(* IEC 61131-3 sources: Elmo_Master/Lasal_PRG/Elmo_EtherCAT_Test_4Axis/Class/CP733_IOs, 1 file *)

(* ---- CP733_IOs.st ---- *)
//FPGA Components
#define CP733_IOS_DEVICE_ID_XADC           16#0A60
#define CP733_IOS_DEVICE_ID_CPU_REG        16#0F02

//XADC Register
#define CP733_IOS_OFFSET_TEMPERATURE       16#00
#define CP733_IOS_OFFSET_VOLTAGE_VP_VN     16#06
#define CP733_IOS_OFFSET_TEMPERATURE_MAX   16#40
#define CP733_IOS_OFFSET_TEMPERATURE_MIN   16#48

//CPU Register
#define CP733_IOS_OFFSET_DIGITAL_INPUT_REGISTER           16#00
#define CP733_IOS_OFFSET_DIGITAL_OUTPUT_CLEAR_REGISTER    16#01
#define CP733_IOS_OFFSET_DIGITAL_OUTPUT_READ_SET_REGISTER 16#02

#define CP733_IOS_REGISTER_NOT_FOUND       16#FFFF

#define CP733_IOS_OFFSET_TEMPSENSOR1       16#08
#define CP733_IOS_OFFSET_TEMPSENSOR2       16#0A

//Constants and calculation from xilinx datasheet
//https://www.xilinx.com/support/documentation/user_guides/ug480_7Series_XADC.pdf
//Equation 2-6 (Temperature) and Equation 2-7 (Voltage)
#define CP733_TEMP_MULTIPLIER    503.975
#define CP733_TEMP_DIVISIOR      4096
#define CP733_TEMP_OFFSET        273.15

#define CP733_IOS_TEMP_CONSTANT_KELVIN  273

#define CP733_VOLTAGE_MULTIPLIER 31

#define CP733_CONVERT_V_TO_MV    1000    //Convert V to mV
#define CP733_CONVERT_TO_1_10_C  10      //Convert °C to 1/10 °C

#define CP733_SUPPLY_VOLTAGE_OFFSET 430  //0,43 V offset (Info from CPU department)

#include "..\..\Source\interfaces\lsl_st_pci.h"
#include "..\..\Source\interfaces\lsl_st_xadc.h"
#include "..\..\Class\PLC_Info\XRegs.h"
#include "..\..\Source\interfaces\lsl_st_gpio.h"

(*!
<Class
	Name               = "CP733_IOs"
	Revision           = "1.0"
	RealtimeTask       = "false"
	CyclicTask         = "false"
	BackgroundTask     = "false"
	Sigmatek           = "true"
	OSInterface        = "false"
	HighPriority       = "false"
	Automatic          = "false"
	UpdateMode         = "Prescan"
	IconPath           = ".\Class\DigInOut.ICO"
	SharedCommandTable = "true"
	Objectsize         = "(688,120)"
	Comment            = "Hardwareclass to access the IOs on the CP733.">
	<Channels>
		<Server Name="BatteryOk" Visualized="true" Initialize="false" WriteProtected="true" Retentive="false" Comment="Shows the state of the battery.&#13;&#10;0 .. Not OK&#13;&#10;1 .. OK"/>
		<Server Name="Can1_Termination" Visualized="true" Initialize="true" WriteProtected="false" Retentive="false" Comment="Write to this server to set the CAN termination.&#13;&#10;0 ... CAN termination is off&#13;&#10;1 ... CAN termination is on&#13;&#10;-1 ... not available/failed to set register in FPGA"/>
		<Server Name="CAN_1_Connect" Class="_CanLib" Visualized="false" Initialize="false" WriteProtected="true" Retentive="false"/>
		<Server Name="ClassState" Visualized="true" Initialize="false" WriteProtected="true" Retentive="false" Comment="Shows the initialisation state of the class.&#13;&#10; 0 ... Initialisation ok&#13;&#10;-1 ... PCI Interface not found&#13;&#10;-2 ... &quot;XADC&quot; interface not found&#13;&#10;-3 ... &quot;IXREGS&quot; interface not found&#13;&#10;-4 ... GPIO Interface not found&#13;&#10;-5 ... CPU Register not found&#13;&#10;-6 ... Login to HwControl failed&#13;&#10;"/>
		<Server Name="ErrorLED" Visualized="true" Initialize="false" WriteProtected="false" Retentive="false" Comment="The &quot;Error&quot;-LED of the CPU can be controlled with this server.&#13;&#10;&#13;&#10;0 ... HW - Status of LED is active&#13;&#10;1 ... LED is off&#13;&#10;2 ... LED is flashes&#13;&#10;3 ... LED is on&#13;&#10;&#13;&#10;-1 ... Class not ok"/>
		<Server Name="Ethernet_1_Connect" Visualized="false" Initialize="false" WriteProtected="true" Retentive="false" Comment="Connection servers for Hardware-Editor."/>
		<Server Name="RunLED" Visualized="true" Initialize="false" WriteProtected="false" Retentive="false" Comment="The &quot;Run&quot;-LED of the CPU can be controlled with this server.&#13;&#10;&#13;&#10;0 ... HW - Status of LED is active&#13;&#10;1 ... LED is off&#13;&#10;2 ... LED is flashes&#13;&#10;3 ... LED is on&#13;&#10;&#13;&#10;-1 ... Class not ok"/>
		<Server Name="StatusLED" Visualized="true" Initialize="false" WriteProtected="false" Retentive="false" Comment="The &quot;Status&quot;-LED of the CPU can be controlled with this server.&#13;&#10;&#13;&#10;0 ... HW - Status of LED is active&#13;&#10;1 ... LED is off&#13;&#10;2 ... LED is flashes&#13;&#10;3 ... LED is on&#13;&#10;&#13;&#10;-1 ... Class not ok"/>
		<Server Name="SupplyVoltage" Visualized="true" Initialize="false" WriteProtected="true" Retentive="false" Comment="Shows the supply voltage in mV."/>
		<Server Name="TemperatureConnectors" Visualized="true" Initialize="false" WriteProtected="true" Retentive="false" Comment="Shows the measured ambient temperature of the connectors in [1°C/10]."/>
		<Server Name="TemperatureCPU" Visualized="true" Initialize="false" WriteProtected="true" Retentive="false" Comment="Shows the measured ambient temperature of the CPU in [1°C/10]."/>
		<Server Name="USB_1_Connect" Visualized="false" Initialize="false" WriteProtected="true" Retentive="false"/>
		<Client Name="To_HwControl" Required="true" Internal="false" Comment="Connect this client to the class &quot;HwControl&quot;."/>
		<Client Name="XXXBase_IOs6" Required="true" Internal="true"/>
	</Channels>
	<Dependencies>
		<Files>
			<File Path=".\Source\interfaces\lsl_st_pci.h" Include="true"/>
			<File Path=".\Source\interfaces\lsl_st_xadc.h" Include="true"/>
			<File Path=".\Class\PLC_Info\XRegs.h" Include="true"/>
			<File Path=".\Source\interfaces\lsl_st_gpio.h" Include="true"/>
		</Files>
	</Dependencies>
	<RevDoku>
		<Owner Company="Sigmatek" Author="EisMic"/>
		<Dokumentation Revision="1.0" Date="12.12.2019" Author="EisMic" Company="Sigmatek" Description="Initial version."/>
	</RevDoku>
	<Network Name="CP733_IOs">
		<!-- List of Components in this network -->
		<Components>
			<Object
				Name       = "XXXBase_IOs6"
				Class      = "XXXBase_IOs"
				Position   = "(150,120)"
				Visualized = "false">
				<Channels>
					<Server Name="CAN_1_Connect"/>
					<Server Name="CAN_2_Connect"/>
					<Server Name="ClassState"/>
					<Server Name="COM_1_Connect"/>
					<Server Name="COM_2_Connect"/>
					<Server Name="COM_3_Connect"/>
					<Server Name="Ethernet_1_Connect"/>
					<Server Name="Ethernet_2_Connect"/>
					<Server Name="Ethernet_3_Connect"/>
					<Server Name="Ethernet_4_Connect"/>
					<Server Name="USB_1_Connect"/>
					<Client Name="To_HwControl"/>
				</Channels>
			</Object>
		</Components>
		<Comments>
		</Comments>
		<!-- List of Connections in this network -->
		<Connections>
			<Connection Source="this.XXXBase_IOs6" Destination="XXXBase_IOs6.ClassState"/>
			<Connection Source="XXXBase_IOs6.To_HwControl" Destination="this.To_HwControl" Vertices="(150,210),(38,210),"/>
			<Connection Source="this.USB_1_Connect" Destination="XXXBase_IOs6.USB_1_Connect" Vertices="(908,750),(736,270),"/>
			<Connection Source="this.CAN_1_Connect" Destination="XXXBase_IOs6.CAN_1_Connect" Vertices="(908,870),(736,570),"/>
			<Connection Source="this.Ethernet_1_Connect" Destination="XXXBase_IOs6.Ethernet_1_Connect" Vertices="(908,810),(736,330),"/>
		</Connections>
		<!-- Headerfiles -->
		<Options>
		</Options>
	</Network>
</Class>
*)
CP733_IOs : CLASS
  //Servers:
	ClassState 	: SvrChCmd_DINT;
	BatteryOk 	: SvrCh_DINT;
	SupplyVoltage 	: SvrCh_DINT;
	TemperatureConnectors 	: SvrCh_DINT;
	TemperatureCPU 	: SvrCh_DINT;
	RunLED 	: SvrCh_DINT;
	ErrorLED 	: SvrCh_DINT;
	StatusLED 	: SvrCh_DINT;
	Can1_Termination 	: SvrCh_DINT;
	USB_1_Connect 	: SvrChCmd_DINT;
	Ethernet_1_Connect 	: SvrChCmd_DINT;
	CAN_1_Connect 	: SvrChCmd_DINT;
  //Clients:
	To_HwControl 	: CltChCmd_HwControl;
	XXXBase_IOs6 	: CltChCmd_XXXBase_IOs;
  //Variables:
		us_FirstScan 	: USINT;
		p_XADC 	: ^void;
		p_CPUReg 	: ^void;
		pXADC 	: ^LSLAPI_IXADC;
		p_XREGS 	: ^T_XREGS;
		bsLedValue : BSINT
		[
		];

		pGPIO 	: ^LSL_GPIO_TYPE;
		sDigitalOutputReadSetRegisterInfo 	: LSL_LOCALIO_IDINFO;
		sDigitalOutputClearRegisterInfo 	: LSL_LOCALIO_IDINFO;
		udFoundRegisterIndex 	: UDINT;
  //Functions:

	FUNCTION VIRTUAL GLOBAL Init;

	FUNCTION VIRTUAL GLOBAL CyWork
		VAR_INPUT
			EAX 	: UDINT;
		END_VAR
		VAR_OUTPUT
			state (EAX) 	: UDINT;
		END_VAR;

	FUNCTION ConvertVoltage
		VAR_INPUT
			uiVoltage 	: UINT;
			Offset 	: DINT;
		END_VAR
		VAR_OUTPUT
			Voltage 	: DINT;
		END_VAR;

	FUNCTION VIRTUAL GLOBAL RunLED::Write
		VAR_INPUT
			input (EAX) 	: DINT;
		END_VAR
		VAR_OUTPUT
			result (EAX) 	: DINT;
		END_VAR;

	FUNCTION VIRTUAL GLOBAL ErrorLED::Write
		VAR_INPUT
			input (EAX) 	: DINT;
		END_VAR
		VAR_OUTPUT
			result (EAX) 	: DINT;
		END_VAR;

	FUNCTION VIRTUAL GLOBAL StatusLED::Write
		VAR_INPUT
			input (EAX) 	: DINT;
		END_VAR
		VAR_OUTPUT
			result (EAX) 	: DINT;
		END_VAR;

	FUNCTION VIRTUAL GLOBAL Can1_Termination::Write
		VAR_INPUT
			input (EAX) 	: DINT;
		END_VAR
		VAR_OUTPUT
			result (EAX) 	: DINT;
		END_VAR;

	FUNCTION VIRTUAL GLOBAL USB_1_Connect::Read
		VAR_OUTPUT
			output (EAX) 	: DINT;
		END_VAR;

	FUNCTION VIRTUAL GLOBAL Ethernet_1_Connect::Read
		VAR_OUTPUT
			output (EAX) 	: DINT;
		END_VAR;

	FUNCTION VIRTUAL GLOBAL CAN_1_Connect::Read
		VAR_OUTPUT
			output (EAX) 	: DINT;
		END_VAR;
  //Tables:
	FUNCTION @STD
		VAR_OUTPUT
			ret_code	: CONFSTATES;
		END_VAR;
	FUNCTION GLOBAL TAB @CT_;
END_CLASS;

#pragma using XXXBase_IOs
#pragma usingLtd HwControl

FUNCTION VIRTUAL GLOBAL CP733_IOs::Init
  VAR
    SigmaTekDevInfo     : ^PCICONFDATA;
    pSPCIInfo           : ^LSL_SPCIINFO;
    Settings            : t_HwObjListSettings;
    result              : DINT;
    tmpLocalIOInfo      : LSL_LOCALIO_IDINFO;
    udAmountLocalIOs    : UDINT;
    i                   : UDINT;
  END_VAR

  us_FirstScan += 1; //Init-counter

  if us_FirstScan = 10 then

    if OS_CILGET("PCICONFIG", #pSPCIInfo) <> SYS_ERR_NONE then
      ClassState := -1; //PCICONFIG not found
      return;
    end_if;

    if OS_CILGET(INTERFACE_XADC, #pXADC) <> SYS_ERR_NONE then
      ClassState := -2; //XADC Device not found
      return;
    end_if;

    if OS_CILGET("IXREGS", #p_XREGS) <> SYS_ERR_NONE then
      ClassState := -3; //XREGS Device not found
      return;
    end_if;

    if OS_CILGET(INTERFACE_GPIO, #pGPIO) <> SYS_ERR_NONE then
      ClassState := -4; //GPIO Device not found
      return;
    end_if;

    SigmaTekDevInfo := SPCIINFO_FINDDEVICE(CP733_IOS_DEVICE_ID_CPU_REG,0);

    //Check pointer to be valid
    if SigmaTekDevInfo then

      p_CPUReg$pVoid := SPCIINFO_GETADDRESS(SigmaTekDevInfo);

      //Check pointer to be valid
      if p_CPUReg = NIL then
        ClassState := 5;
        return;
      end_if;
    else
      ClassState := -5;
      return;
    end_if;

    //Get necessary infos for Can termination handling
    //*********************************************************************************************************************

    //Get amount of local IOs from OS
    udAmountLocalIOs      := OS_LOCALIO_GETCOUNT(pGPIO);
    udFoundRegisterIndex  := CP733_IOS_REGISTER_NOT_FOUND; //Register not found

    //Check if we found local IOs on the hardware
    if udAmountLocalIOs then

      //Now search all local IOs to find the correct registers of the "wb_cpu_reg" component
      for i:= 0 to udAmountLocalIOs-1 do
        result := OS_LOCALIO_GETINFO(pGPIO,i,#tmpLocalIOInfo);

        //Check if we found the correct component
        if (tmpLocalIOInfo.typeinfo AND 16#FFFF) = CP733_IOS_DEVICE_ID_CPU_REG then

          //We found it, save number and exit
          udFoundRegisterIndex := i;
          exit;
        end_if;
      end_for;

      //Check if we found the correct component
      if udFoundRegisterIndex <> CP733_IOS_REGISTER_NOT_FOUND then

        //Now we have to get the correct ID of both the "Clear" and the "Read/Set" Register
        //First local io we found is the Digital Input Reg because it is the first one in the adress mapping

        //Reg 0 ... Digital Input               ... udFoundRegisterIndex
        //Reg 1 ... Digtal Output Clear         ... udFoundRegisterIndex + 1
        //Reg 2 ... Digital Output Read / Set   ... udFoundRegisterIndex + 2

        result := OS_LOCALIO_GETINFO(pGPIO,udFoundRegisterIndex + CP733_IOS_OFFSET_DIGITAL_OUTPUT_CLEAR_REGISTER,#sDigitalOutputClearRegisterInfo);

        //Check for errors
        if result <> 0 then
          udFoundRegisterIndex  := CP733_IOS_REGISTER_NOT_FOUND; //Register not found
        end_if;

        result := OS_LOCALIO_GETINFO(pGPIO,udFoundRegisterIndex + CP733_IOS_OFFSET_DIGITAL_OUTPUT_READ_SET_REGISTER,#sDigitalOutputReadSetRegisterInfo);

        //Check for errors
        if result <> 0 then
          udFoundRegisterIndex  := CP733_IOS_REGISTER_NOT_FOUND; //Register not found
        end_if;
      end_if;
    end_if;

    //Write first time in init
    Can1_Termination.Write(input:=Can1_Termination);

    //*********************************************************************************************************************

    // initialisiation OK => we login to HwControl
    Settings            := 0;
    Settings.Cyclic     := TRUE;

    if To_HwControl.AddHwObject(pThis:=THIS$pVirtualBase, Settings:=Settings) then
      ClassState := -6;
    end_if;
  end_if;

END_FUNCTION

FUNCTION VIRTUAL GLOBAL CP733_IOs::CyWork
	VAR_INPUT
		EAX 	: UDINT;
	END_VAR
	VAR_OUTPUT
		state (EAX) 	: UDINT;
	END_VAR
  VAR
  	udTmpValue : UDINT;
  END_VAR

  //Check if initialisation was successfull -> so pointers must be valid and we don't need to check them
  if ClassState = 0 then

    OS_XADC_GETVPVN(pXADC,#udTmpValue);
    SupplyVoltage           := ConvertVoltage(udTmpValue$UINT,CP733_SUPPLY_VOLTAGE_OFFSET);

    TemperatureConnectors   := ((p_CPUReg + 16#8)^$UINT - CP733_IOS_TEMP_CONSTANT_KELVIN) * CP733_CONVERT_TO_1_10_C;
    TemperatureCPU          := ((p_CPUReg + 16#A)^$UINT - CP733_IOS_TEMP_CONSTANT_KELVIN) * CP733_CONVERT_TO_1_10_C;

    BatteryOk := p_XREGS^.Batt_funct$funct_XREGS_BattGood();

  else
    //Show on server that the information is not valid
    SupplyVoltage           := ACCESS_DENIED;
    TemperatureConnectors   := ACCESS_DENIED;
    TemperatureCPU          := ACCESS_DENIED;
    RunLED                  := -1;
    ErrorLED                := -1;
    StatusLED               := -1;
  end_if;

	state := READY;

END_FUNCTION

FUNCTION CP733_IOs::ConvertVoltage
	VAR_INPUT
		uiVoltage 	: UINT;
		Offset 	: DINT;
	END_VAR
	VAR_OUTPUT
		Voltage 	: DINT;
	END_VAR

  //12 Bit Value is stored in the MSB bits in the 16bit register -> shift right 4
  Voltage := TO_DINT( TO_REAL(((uiVoltage SHR 4) * CP733_VOLTAGE_MULTIPLIER * CP733_CONVERT_V_TO_MV) / CP733_TEMP_DIVISIOR));
  Voltage += Offset;

END_FUNCTION

FUNCTION VIRTUAL GLOBAL CP733_IOs::RunLED::Write
	VAR_INPUT
		input (EAX) 	: DINT;
	END_VAR
	VAR_OUTPUT
		result (EAX) 	: DINT;
	END_VAR

  if p_XREGS then
    if input >= 0 & input <= 3 then
      RunLED := input;
      bsLedValue := (RunLED$USINT AND 0x3) OR ((StatusLED$USINT AND 0x3) SHL 2) OR ((ErrorLED$USINT AND 0x3) SHL 4);
      p_XREGS^.LED_funct$funct_XREGS_SETLeds(val:= bsLedValue);
    end_if;
  end_if;

	result := RunLED;

END_FUNCTION

FUNCTION VIRTUAL GLOBAL CP733_IOs::ErrorLED::Write
	VAR_INPUT
		input (EAX) 	: DINT;
	END_VAR
	VAR_OUTPUT
		result (EAX) 	: DINT;
	END_VAR

  if p_XREGS then
    if input >= 0 & input <= 3 then
      ErrorLED := input;
      bsLedValue := (RunLED$USINT AND 0x3) OR ((StatusLED$USINT AND 0x3) SHL 2) OR ((ErrorLED$USINT AND 0x3) SHL 4);
      p_XREGS^.LED_funct$funct_XREGS_SETLeds(val:= bsLedValue);
    end_if;
  end_if;

	result := ErrorLED;

END_FUNCTION

FUNCTION VIRTUAL GLOBAL CP733_IOs::StatusLED::Write
	VAR_INPUT
		input (EAX) 	: DINT;
	END_VAR
	VAR_OUTPUT
		result (EAX) 	: DINT;
	END_VAR

  if p_XREGS then
    if input >= 0 & input <= 3 then
      StatusLED := input;
      bsLedValue := (RunLED$USINT AND 0x3) OR ((StatusLED$USINT AND 0x3) SHL 2) OR ((ErrorLED$USINT AND 0x3) SHL 4);
      p_XREGS^.LED_funct$funct_XREGS_SETLeds(val:= bsLedValue);
    end_if;
  end_if;

	result := StatusLED;

END_FUNCTION

FUNCTION VIRTUAL GLOBAL CP733_IOs::Can1_Termination::Write
	VAR_INPUT
		input (EAX) 	: DINT;
	END_VAR
	VAR_OUTPUT
		result (EAX) 	: DINT;
	END_VAR
  VAR
    TmpRegValue : UDINT;
  END_VAR

  //Digitale Ausgänge
  //Bit 0: USB 0 einschalten (wird noch nicht verwendet)
  //Bit 1: USB 3.0 einschalten(wird noch nicht verwendet)
  //Bit 2: USB 2 einschalten(wird noch nicht verwendet)
  //Bit 3: USB 3 einschalten(wird noch nicht verwendet)
  //Bit 4: CPU Power BTN
  //Bit 5: Can TERM einschalten
  //Bit 6: SDIAS 24V einschalten
  //Bit 7: SDIAS 5V einschalten
  //Bit 15..8: Reserviert

  //Check if function is available
  if pGPIO & udFoundRegisterIndex <> CP733_IOS_REGISTER_NOT_FOUND then

    //Get current register value
    result$DINT := OS_GPIO_GETREG(pGPIO, sDigitalOutputReadSetRegisterInfo.id, CP733_IOS_OFFSET_DIGITAL_OUTPUT_READ_SET_REGISTER, #TmpRegValue);

    //Check for errors
    if result = 0 then

      //Register in FPGA is inverted
      //*****************************************************************************
      if input = 1 then

        TmpRegValue := 0x20;  //Only clear Bit 5

        result$DINT := OS_GPIO_SETREG(pGPIO, sDigitalOutputClearRegisterInfo.id, CP733_IOS_OFFSET_DIGITAL_OUTPUT_CLEAR_REGISTER, TmpRegValue);

        if result = 0 then
          Can1_Termination := 1;
        else
          Can1_Termination := -1; //Failed to set register
        end_if;

      //*****************************************************************************
      elsif input = 0 then

        TmpRegValue := TmpRegValue OR 0x20;  //Set current Bits and Bit 5

        result$DINT := OS_GPIO_SETREG(pGPIO, sDigitalOutputReadSetRegisterInfo.id, CP733_IOS_OFFSET_DIGITAL_OUTPUT_READ_SET_REGISTER, TmpRegValue);

        if result = 0 then
          Can1_Termination := 0;
        else
          Can1_Termination := -1; //Failed to set register
        end_if;
      end_if;
      //*****************************************************************************
    else
      Can1_Termination := -1;
    end_if;
  else
    Can1_Termination := -1;
  end_if;

	result := Can1_Termination;

END_FUNCTION

FUNCTION VIRTUAL GLOBAL CP733_IOs::USB_1_Connect::Read
	VAR_OUTPUT
		output (EAX) 	: DINT;
	END_VAR

	USB_1_Connect := XXXBase_IOs6.USB_1_Connect.Read();
	output := USB_1_Connect;

END_FUNCTION

FUNCTION VIRTUAL GLOBAL CP733_IOs::CAN_1_Connect::Read
	VAR_OUTPUT
		output (EAX) 	: DINT;
	END_VAR

	CAN_1_Connect := XXXBase_IOs6.CAN_1_Connect.Read();
	output := CAN_1_Connect;

END_FUNCTION

FUNCTION VIRTUAL GLOBAL CP733_IOs::Ethernet_1_Connect::Read
	VAR_OUTPUT
		output (EAX) 	: DINT;
	END_VAR

	Ethernet_1_Connect := XXXBase_IOs6.Ethernet_1_Connect.Read();
	output := Ethernet_1_Connect;

END_FUNCTION
